Staubli VAL3: Lab2B_L3.pjx

--- Lab2B_L3.pjx ---
parameters version=s6.8 stackSize=5000 millimeterUnit=true
program file=start.pgx
program file=feedCylinder.pgx
program file=placeCylinder.pgx
program file=insertPiston.pgx
program file=placeInMatrix.pgx
program file=physicalIO.pgx
program file=stop.pgx
data file=Lab2B_L3.dtx
alias name=io interface=io autoload=true

--- Lab2B_L3.dtx ---


--- start.pgx ---
program start()
// Level 3: four taught piston slots with tool presence sensing and bounded assembly.
  local num poseIndex
  local point approachPose
  local point placePose
  local point pistonApproach
  local point pickPose
  local point checkPose
  local point checkApproach
begin
  // ============================================================
  // LEVEL 3: ALIMENTAR, MONTAR Y COLOCAR CUATRO CONJUNTOS
  // ============================================================
  // Adaptacion Level 2 de la estructura de Isma; originales preservados.
  // Lab2B (Level 1) y Lab2B_Level2 permanecen sin modificar.
  // Matriz VACIA. Los huecos sin piston se detectan y se omiten.
  // simulation=true: sensores manuales, sin acceso a pines.
  // simulation=false: bIn2/14/15, bOut10 y pinza valve1.
  userPage()
  cls()
  putln("Lab2B_L3 - Four assemblies - empty matrix required")
  physicalRun = !simulation
  placedCount = 0
  partIndex = 0
  pistonIndex = 0
  pistonFound = false
  pistonChecked = false
  cycleStep = 0
  feederExtend = false
  ioReady = false

  // ============================================================
  // COMPROBAR ALTURAS DE MATRIZ SIN MOVER NI ACCIONAR SALIDAS
  // ============================================================
  // Parejas 0/1, 2/3, 4/5, 6/7: par=approach, impar=deposito.
  // J3 es un ANGULO, no una altura. Calculamos Z del TCP lateral.
  // Esto comprueba altura, no colisiones, alineacion o alcance del trayecto.
  for poseIndex = 0 to 3
    approachPose = jointToPoint(tLateral, world, jMatrix[2*poseIndex])
    placePose = jointToPoint(tLateral, world, jMatrix[2*poseIndex+1])
    putln("Matrix slot (0..3):")
    putln(poseIndex)
    putln("Approach Z (mm):")
    putln(approachPose.trsf.z)
    putln("Place Z (mm):")
    putln(placePose.trsf.z)
    if approachPose.trsf.z <= placePose.trsf.z
      putln("ERROR: approach is not above place; review this matrix pair")
      return
    endIf
  endFor

  // ============================================================
  // CUATRO RECOGIDAS REALES: IMG_3805, 3806, 3807, 3808
  // ============================================================
  // jPistonPick: impares = recogidas ENSENADAS; pares = approaches
  // CALCULADOS aqui (pick + pistonLift en Z world, misma orientacion).
  // jPistonCheck[0..3]: poses de deteccion bIn0 ENSENADAS en el mando
  // (sensor lateral de la pinza). NO se recalculan ni se sobrescriben.
  // jCheckApproach[0..3]: CALCULADOS aqui (check + checkLift en Z world,
  // misma orientacion). Los ceros del DTX son espacio para el resultado.
  // Todo termina antes de crear tareas o mover el robot.
  if pistonLift <= 0 or checkLift <= 0
    putln("ERROR: pistonLift and checkLift must be positive (mm)")
    return
  endIf
  for poseIndex = 0 to 3
    if jPistonPick[2*poseIndex+1].j1 == 0 and jPistonPick[2*poseIndex+1].j2 == 0 and jPistonPick[2*poseIndex+1].j3 == 0 and jPistonPick[2*poseIndex+1].j4 == 0 and jPistonPick[2*poseIndex+1].j5 == 0 and jPistonPick[2*poseIndex+1].j6 == 0
      putln("ERROR: teach piston pick joint; missing piston (0..3):")
      putln(poseIndex)
      return
    endIf
    if jPistonCheck[poseIndex].j1 == 0 and jPistonCheck[poseIndex].j2 == 0 and jPistonCheck[poseIndex].j3 == 0 and jPistonCheck[poseIndex].j4 == 0 and jPistonCheck[poseIndex].j5 == 0 and jPistonCheck[poseIndex].j6 == 0
      putln("ERROR: teach jPistonCheck; missing sensing pose (0..3):")
      putln(poseIndex)
      return
    endIf
    pickPose = jointToPoint(tTip, world, jPistonPick[2*poseIndex+1])
    pistonApproach = pickPose
    pistonApproach.trsf.z = pickPose.trsf.z + pistonLift
    if !pointToJoint(tTip, jPistonPick[2*poseIndex+1], pistonApproach, jPistonPick[2*poseIndex])
      putln("ERROR: no piston approach solution; piston (0..3):")
      putln(poseIndex)
      return
    endIf
    checkPose = jointToPoint(tTip, world, jPistonCheck[poseIndex])
    checkApproach = checkPose
    checkApproach.trsf.z = checkPose.trsf.z + checkLift
    if !pointToJoint(tTip, jPistonCheck[poseIndex], checkApproach, jCheckApproach[poseIndex])
      putln("ERROR: no check approach solution; piston (0..3):")
      putln(poseIndex)
      return
    endIf
    putln("Piston slot (0..3):")
    putln(poseIndex)
    putln("  tTip Z pick / pickAppr / check / checkAppr (mm):")
    putln(pickPose.trsf.z)
    putln(pistonApproach.trsf.z)
    putln(checkPose.trsf.z)
    putln(checkApproach.trsf.z)
    putln("  check - pick XY offset (mm):")
    putln(checkPose.trsf.x - pickPose.trsf.x)
    putln(checkPose.trsf.y - pickPose.trsf.y)
  endFor

  // physicalIO solo escribe el ALIMENTADOR; nunca la pinza.
  if physicalRun
    taskCreate "physicalIO", 10, physicalIO()
    wait(ioReady == true)
    putln("PHYSICAL: real sensors and feeder enabled")
    open(tLateral)
  else
    putln("MANUAL SIMULATION: change sensor bools at the indicated steps")
    delay(tLateral.otime)
  endIf
  movej(jStart[0], tLateral, mNomSpeed)
  waitEndMove()

  // ============================================================
  // SOLO CUATRO CONJUNTOS; NO HAY QUINTA ALIMENTACION
  // ============================================================
  while placedCount < 4
    partIndex = placedCount
    putln("Assembly number (1..4):")
    putln(partIndex+1)
    call feedCylinder()
    call placeCylinder()
    call insertPiston()
    call placeInMatrix()
    // Contar tras soltar y terminar la retirada de la matriz.
    placedCount = placedCount + 1
    putln("Completed matrix slots:")
    putln(placedCount)
    // Volver a la postura inicial SOLO si falta otro conjunto.
    if placedCount < 4
      movej(jStart[0], tLateral, mNomSpeed)
      waitEndMove()
    endIf
  endWhile

  // La matriz llena finaliza aunque bIn2 siga detectando cilindros.
  feederExtend = false
  taskKill("physicalIO")
  if physicalRun
    io:bOut10 = false
  endIf
  ioReady = false
  cycleStep = 100
  putln("100 - Matrix full: 4/4. No further feeding or pickup.")
end

--- feedCylinder.pgx ---
program feedCylinder()
// Level 3: four taught piston slots with tool presence sensing and bounded assembly.
begin
  // ============================================================
  // PREPARAR UN CILINDRO, CON EL ROBOT FUERA DEL DISPENSADOR
  // ============================================================
  // bOut10: 1=extender, 0=retraer (mapa del enunciado).
  // bIn14/bIn15: finales extendido/retraido; bIn2: cilindro listo.
  // El PDF no especifica toda la secuencia mecanica: se propone
  // extender y retraer antes de entrar con el robot. Verificar en la celda.
  // Si ya hay un cilindro preparado, no empujar otro encima.
  cycleStep = 10
  feederExtend = false
  putln("10 - Wait feederRetracted=true and feederExtended=false")
  wait(feederRetracted == true and feederExtended == false)
  if !cylinderPresent
    cycleStep = 11
    putln("11 - EXTEND feeder; wait extended=true / retracted=false")
    feederExtend = true
    wait(feederExtended == true and feederRetracted == false)

    cycleStep = 12
    putln("12 - RETRACT feeder; wait retracted=true / extended=false")
    feederExtend = false
    wait(feederRetracted == true and feederExtended == false)
  endIf
  cycleStep = 13
  putln("13 - Wait cylinderPresent=true; cylinder ready for pickup")
  wait(cylinderPresent == true)
end

--- insertPiston.pgx ---
program insertPiston()
// Level 3: four taught piston slots with tool presence sensing and bounded assembly.
begin
  // ============================================================
  // 40-43. BUSCAR UN PISTON: REVISAR SIEMPRE LOS 4 HUECOS DESDE EL 0
  // ============================================================
  // En cada montaje se recorre pistonIndex = 0,1,2,3 y se coge el
  // PRIMER hueco donde bIn0 detecta piston. partIndex solo cuenta montajes.
  // bIn0 esta en un LATERAL de la pinza y detecta presencia, no agarre.
  // Por hueco (todo con tTip):
  //   40 movej jCheckApproach (check + checkLift, calculado en start)
  //      movel jPistonCheck (ENSENADA) -> 41 leer bIn0
  //   Si NO hay piston: no se retira; se va directo al siguiente hueco.
  //   Si hay piston: 42 subir a jCheckApproach, ir al approach del pick,
  //      bajar vertical a jPistonPick, cerrar y subir al approach.
  // Si los 4 estan vacios: subir, avisar, esperar 2 s y repetir desde 0.
  pistonFound = false
  if physicalRun
    open(tTip)
  else
    delay(tTip.otime)
  endIf
  while !pistonFound
    pistonIndex = 0
    while !pistonFound and pistonIndex < 4
      cycleStep = 40
      putln("40 - Check piston slot (0..3):")
      putln(pistonIndex)
      putln("DBG 40A - movej to check approach")
      movej(jCheckApproach[pistonIndex], tTip, mNomSpeed)
      waitEndMove()
      putln("DBG 40B - movel to taught sensing pose jPistonCheck")
      movel(jointToPoint(tTip, world, jPistonCheck[pistonIndex]), tTip, mApproachSpeed)
      waitEndMove()
      cycleStep = 41
      pistonChecked = false
      if physicalRun
        // Asentar la herramienta y dejar actualizar physicalIO antes de leer.
        delay(0.15)
      else
        putln("MANUAL: set pistonPresent, then pistonChecked=true")
        wait(pistonChecked == true)
      endIf
      // Guardar la lectura ANTES de mover: physicalIO sigue refrescando
      // pistonPresent y al alejarse el sensor dejaria de verlo.
      pistonFound = pistonPresent
      putln("41 - Tool presence sensor bIn0:")
      if pistonFound
        putln("pistonPresent = true")
      else
        putln("pistonPresent = false")
        cycleStep = 43
        putln("43 - Empty slot; go to next slot")
        pistonIndex = pistonIndex + 1
      endIf
    endWhile
    if !pistonFound
      // Ultimo check fue el hueco 3: subir antes de volver al hueco 0.
      movel(jointToPoint(tTip, world, jCheckApproach[3]), tTip, mApproachSpeed)
      waitEndMove()
      putln("No piston in any slot; refill tray. Rescanning in 2 s.")
      delay(2)
    endIf
  endWhile

  // pistonIndex = primer hueco con piston detectado.
  cycleStep = 42
  putln("42 - Piston found; pick slot (0..3):")
  putln(pistonIndex)
  putln("DBG 42A - movel up to check approach")
  movel(jointToPoint(tTip, world, jCheckApproach[pistonIndex]), tTip, mApproachSpeed)
  waitEndMove()
  putln("DBG 42B - movel to pick approach")
  movel(jointToPoint(tTip, world, jPistonPick[2*pistonIndex]), tTip, mApproachSpeed)
  waitEndMove()
  putln("DBG 42C - movel down to pick; then close tTip")
  movel(jointToPoint(tTip, world, jPistonPick[2*pistonIndex+1]), tTip, mApproachSpeed)
  waitEndMove()
  if physicalRun
    close(tTip)
  else
    delay(tTip.ctime)
  endIf
  putln("DBG 42D - Piston gripped; withdraw to pick approach")
  movel(jointToPoint(tTip, world, jPistonPick[2*pistonIndex]), tTip, mApproachSpeed)
  waitEndMove()

  // ============================================================
  // 50. INSERTAR EL PISTON Y SOLTARLO ANTES DE RETIRARSE
  // ============================================================
  // TODO SIMULACION: confirmar el orden [0]/[1] de gridpiston.
  // TODO FISICO: ajustar alineacion y profundidad de jPistonInsert[1].
  // Este movimiento es por posicion; no mide fuerza ni confirma montaje.
  cycleStep = 50
  putln("50 - Insert piston into cylinder")
  putln("DBG 50A - BEFORE movej: insertion approach [0]")
  movej(jPistonInsert[0], tTip, mNomSpeed)
  waitEndMove()
  putln("DBG 50B - Insertion approach reached")
  movej(jointToPoint(tTip, world, jPistonInsert[1]), tTip, mInsertSpeed)
  waitEndMove()
  putln("DBG 50C - Insertion reached with tTip; opening gripper")
  if physicalRun
    open(tTip)
  else
    delay(tTip.otime)
  endIf
  putln("DBG 50D - BEFORE withdrawal with tTip to jPistonInsert[0]")
  movej(jointToPoint(tTip, world, jPistonInsert[0]), tTip, mInsertSpeed)
  waitEndMove()
  putln("DBG 50E - Tip withdrawal completed")

  // ============================================================
  // 55. POSTURA INTERMEDIA ANTES DE RECOGER EL CONJUNTO
  // ============================================================
  // Joint indicada por el usuario. Se alcanza DESPUES de soltar
  // el piston y retirarse con tTip, antes del agarre con tLateral.
  cycleStep = 55
  putln("DBG 55A - BEFORE movej: jAssemblyMove with tTip")
  movej(jAssemblyMove, tTip, mNomSpeed)
  waitEndMove()
  putln("DBG 55B - Assembly transit posture reached")

end

--- physicalIO.pgx ---
program physicalIO()
// Level 3: four taught piston slots with tool presence sensing and bounded assembly.
begin
  // ============================================================
  // SENSORES Y ALIMENTADOR DEL LEVEL 3
  // ============================================================
  // Solo se crea en fisico. En simulacion los sensores se editan a mano.
  // La pinza usa open/close con valve1; NO escribir valve1 aqui.
  while true
    pistonPresent = io:bIn0 == true
    cylinderPresent = io:bIn2 == true
    feederExtended = io:bIn14 == true
    feederRetracted = io:bIn15 == true
    io:bOut10 = feederExtend
    ioReady = true
    delay(0.01)
  endWhile
end

--- placeCylinder.pgx ---
program placeCylinder()
// Level 3: four taught piston slots with tool presence sensing and bounded assembly.
begin
  // partIndex=0..3 selecciona la pareja del piston correspondiente.
  // ============================================================
  // 20. RECOGER EL CILINDRO CON EL TCP LATERAL
  // ============================================================
  // movej: traslado articular entre aproximaciones.
  // movel: entradas/retiradas con mApproachSpeed; insercion con mInsertSpeed.
  // jointToPoint convierte la joint para movel; no mueve el robot.
  // Usar el mismo TCP en la conversion y en la orden de movimiento.
  // waitEndMove termina cada movimiento antes de accionar la pinza.
  cycleStep = 20
  putln("20 - Pick cylinder - tLateral")
  movej(jCylinderPick[0], tLateral, mNomSpeed)
  waitEndMove()
  movel(jointToPoint(tLateral, world, jCylinderPick[1]), tLateral, mApproachSpeed)
  waitEndMove()

  // Cerrar y dar el tiempo mecanico guardado en la herramienta (1 s).
  // No hay confirmacion de agarre en el mapa de E/S de esta practica.
  if physicalRun
    close(tLateral)
  else
    delay(tLateral.ctime)
  endIf
  movel(jointToPoint(tLateral, world, jCylinderPick[0]), tLateral, mApproachSpeed)
  waitEndMove()
  // El cilindro ya se ha retirado: exigir sensor libre antes
  // de admitir otra alimentacion en la siguiente vuelta.
  cycleStep = 21
  putln("21 - Wait cylinderPresent=false after cylinder withdrawal")
  wait(cylinderPresent == false)

  // ============================================================
  // 30. DEPOSITAR EL CILINDRO EN LA ESTACION DE MONTAJE
  // ============================================================
  cycleStep = 30
  putln("30 - Place cylinder at assembly station")
  movej(jCylinderPlace[0], tLateral, mNomSpeed)
  waitEndMove()
  movel(jointToPoint(tLateral, world, jCylinderPlace[1]), tLateral, mApproachSpeed)
  waitEndMove()
  if physicalRun
    open(tLateral)
  else
    delay(tLateral.otime)
  endIf
  movel(jointToPoint(tLateral, world, jCylinderPlace[0]), tLateral, mApproachSpeed)
  waitEndMove()

end

--- placeInMatrix.pgx ---
program placeInMatrix()
// Level 3: four taught piston slots with tool presence sensing and bounded assembly.
begin
  // ============================================================
  // 60. RECOGER EL CONJUNTO CON EL TCP LATERAL
  // ============================================================
  // Recoger en jCylinderPlace[1], donde se ha depositado el cilindro.
  // TODO FISICO: comprobar el agarre con el piston ya dentro del cilindro.
  cycleStep = 60
  putln("60 - Pick assembled cylinder - tLateral")
  if physicalRun
    open(tLateral)
  else
    delay(tLateral.otime)
  endIf
  // El siguiente movimiento usa el TCP lateral. Las joints guardadas
  // deben describir la postura de agarre lateral; el TCP no anade un giro.
  putln("DBG 60A - BEFORE movej with tLateral to jCylinderPlace[0]")
  movej(jCylinderPlace[0], tLateral, mNomSpeed)
  waitEndMove()
  putln("DBG 60B - Lateral approach reached; BEFORE descent to jCylinderPlace[1]")
  movel(jointToPoint(tLateral, world, jCylinderPlace[1]), tLateral, mApproachSpeed)
  waitEndMove()
  putln("DBG 60C - Assembly pickup reached with tLateral; closing gripper")
  if physicalRun
    close(tLateral)
  else
    delay(tLateral.ctime)
  endIf
  putln("DBG 60D - BEFORE withdrawal of assembly with tLateral")
  movel(jointToPoint(tLateral, world, jCylinderPlace[0]), tLateral, mApproachSpeed)
  waitEndMove()
  putln("DBG 60E - Assembly withdrawal completed")

  // ============================================================
  // DEPOSITAR EN LA PAREJA DEL HUECO ACTUAL DE LA MATRIZ
  // ============================================================
  // partIndex es 0..3: approach=2*i, deposito=2*i+1.
  // El llamador limita a cuatro y pasa el indice correspondiente.
  cycleStep = 70
  putln("70 - Place assembly in matrix slot (0..3):")
  putln(partIndex)
  movej(jMatrix[2*partIndex], tLateral, mNomSpeed)
  waitEndMove()
  movel(jointToPoint(tLateral, world, jMatrix[2*partIndex+1]), tLateral, mApproachSpeed)
  waitEndMove()
  if physicalRun
    open(tLateral)
  else
    delay(tLateral.otime)
  endIf
  movel(jointToPoint(tLateral, world, jMatrix[2*partIndex]), tLateral, mApproachSpeed)
  waitEndMove()
  putln("75 - Assembly released; matrix withdrawal completed")
end

--- stop.pgx ---
program stop()
// Level 3: four taught piston slots with tool presence sensing and bounded assembly.
begin
  // Detener el adaptador antes de mandar retraer el alimentador.
  // taskKill no hace nada si la tarea no existe (p. ej. setup incompleto).
  taskKill("physicalIO")
  resetMotion()
  feederExtend = false
  // No tocar hardware si start termino por posiciones pendientes.
  if physicalRun and ioReady
    io:bOut10 = false
  endIf
  ioReady = false
  cycleStep = -1
  // No abrir/cerrar la pinza ni ordenar retorno automatico.
  // Un nuevo start reinicia el contador: vaciar matriz antes de reiniciar.
  putln("STOP - Feeder retract command; gripper unchanged. Prepare cell before restart.")
end
